(* IEC 61131-3 sources: daoli-st-library/DL_Device (part 37) *)

(* ---- FB_DL_WaferCassetteSlot.st ---- *)
(*==============================================================================
 * 组件名称 (Component)  : FB_DL_WaferCassetteSlot
 * 所属子库 (Sublibrary) : DL_Device
 * 当前版本 (Version)    : 1.0.0
 * 兼容性 (Platform)     : CODESYS 3.5 / TwinCAT 3 / 汇川 InoProShop（纯标准元素，零方言）
 * 功能描述 (Function)   : 花篮 25 槽占用双向计数与满/空判据。进片沿 +1、出片沿 −1，同拍
 *                         双沿按「物理不可能，必是抖动或逻辑错」双丢弃并报码；两个沿的净
 *                         额一次性施加，占用计数只有一处写入点；占用为 0 时的出片不借位到
 *                         25（借位会把满篮误判为空篮），锁存计数矛盾；位图按先低槽后高槽
 *                         顺序填充（顺序装片假设），出片清最低置位位。不做槽位光学检测、
 *                         不做花篮身份识别。
 * 溯源 (Origin)         : 道莅 clean-room 防御性实现
 * 本文件内含 (Contains) : TYPE E_DL_CassetteState / FUNCTION_BLOCK FB_DL_WaferCassetteSlot
 * 依赖 (Depends)        : 无（仅 Standard.library 的 SHL / SHR 与位运算）
 * 红线自检 (Redline)    : 无外部全局变量、无硬件地址直引 ｜ 全变量中英双语同行注释
 *                         槽数钳位 1~25 且写位图前判槽号 ｜ 占用计数单点写入（净额合并）
 *                         双沿沿实例无条件周期刷新 ｜ 枚举显式赋值 ｜ CASE 含 ELSE 兜底
 * 错误码表 (Codes)      : 16#0003_03B6 就绪（计数正常，含满/空稳态）
 *                         16#0003_03B7 故障级 清空请求在使能期被拒（清空须先失能）
 *                         16#0003_03B8 信息级 槽数 >25 已钳制（不置故障级标志）
 *                         16#0003_03B9 故障级 同拍进出双沿或满篮进片（请求双丢弃）
 *                         16#0003_03BA 故障级 空篮出片，锁存计数矛盾（不借位到 25）。
 *                                    本件 5 槽全用、无预留槽，已登记待裁定
 * 修订历史 (Revision)   : 2026-11-17  v1.0.0  首版入库 · R28 · 阶段三批 3
 * 验收向量 (Acceptance) : 正向 25 槽连续进满 → 占用 25、bFull、位图 16#01FF_FFFF；再出
 *                         1 片 → 占用 24、bFull=FALSE、16#0003_03B6
 *                         反向 空篮出片 → bCounterMismatch、占用保持 0、16#0003_03BA；
 *                         同拍进出双沿 → 16#0003_03B9 且双丢弃；槽数给 30 → 钳 25 +
 *                         16#0003_03B8（信息级）；使能期清空请求 → 16#0003_03B7 且不清
 *============================================================================*)

(*-----------------------------------------------------------------------------
 * 枚举: E_DL_CassetteState（归属本功能块，同文件发布，全库唯一定义）
 *----------------------------------------------------------------------------*)
TYPE E_DL_CassetteState :
(
    eEmpty := 0,    // 空篮：占用 0 / Empty cassette, no occupied slot
    ePart  := 10,   // 部分占用：0 < 占用 < 槽数 / Partially occupied
    eFull  := 20,   // 满篮：占用 = 槽数 / Full cassette
    eFault := 99    // 故障：计数矛盾锁存 / Fault, the counter contradiction is latched
);
END_TYPE

FUNCTION_BLOCK FB_DL_WaferCassetteSlot
VAR_INPUT
    bEnable      : BOOL := FALSE;         // 使能，FALSE 锁存位图（计数冻结） / Enable, FALSE freezes the slot map
    bLoadPulse   : BOOL := FALSE;         // 进片 +1，上升沿 / Load pulse, rising edge adds one
    bUnloadPulse : BOOL := FALSE;         // 出片 −1，上升沿 / Unload pulse, rising edge subtracts one
    bClear       : BOOL := FALSE;         // 清空（换花篮），须 bEnable=FALSE / Clear for a cassette change, requires bEnable FALSE
    uSlotCount   : UINT := 25;            // 槽数 [个]，域 1~25 / Slot count, domain 1 to 25
END_VAR
VAR_OUTPUT
    uOccupied    : UINT;                  // 占用槽数 [个] / Occupied slot count
    uEmptySlot   : UINT;                  // 空槽数 [个] / Empty slot count
    bFull        : BOOL;                  // 满篮判据 / Full criterion
    bEmpty       : BOOL;                  // 空篮判据 / Empty criterion
    uSlotMask    : DWORD;                 // 占用位图 bit0=第 1 槽 … bit24=第 25 槽 [bit]（25 位须 32 位容器，规格 WORD 无法表达） / Occupancy map, 25 bits need a 32-bit container
    bCounterMismatch : BOOL;              // 计数矛盾已锁存 / Counter contradiction latched
    eErr         : UDINT;                 // 错误码，段位 16#0003_xxxx / Error code in segment 16#0003_xxxx
END_VAR
VAR
    _eState      : E_DL_CassetteState := E_DL_CassetteState.eEmpty; // 占用状态 / Occupancy state
    _bInit       : BOOL := FALSE;         // 首扫标志，取非判定 / First-scan flag, tested negated
    _bMismatch   : BOOL := FALSE;         // 矛盾锁存状态量 / Contradiction latch state quantity
    _nNet        : INT;                   // 本拍净额（+进 −出） / Net delta of this scan
    _uSlotEff    : UINT := 25;            // 生效槽数（钳制后） / Effective slot count after clamping
    _uwOccupied  : UINT;                  // 占用内部唯一写点 / The single internal write point of the occupancy
    _rtrigLoad   : R_TRIG;                // 进片上升沿 / Rising edge of the load pulse
    _rtrigUnload : R_TRIG;                // 出片上升沿 / Rising edge of the unload pulse
END_VAR
VAR CONSTANT
    DL_CS_READY   : UDINT := 16#0003_03B6;  // 就绪码 / Ready code
    DL_CS_CLEAR_REJ : UDINT := 16#0003_03B7; // 故障级清空被拒码 / Fault code for a rejected clear request
    DL_CS_SLOT_CLAMP : UDINT := 16#0003_03B8; // 信息级槽数钳制码 / Info code for a clamped slot count
    DL_CS_BOTH    : UDINT := 16#0003_03B9;  // 故障级双沿或满篮进片码 / Fault code for double edges or a load on a full cassette
    DL_CS_UNDER   : UDINT := 16#0003_03BA;  // 故障级空篮出片码 / Fault code for an unload on an empty cassette
    DL_CS_SLOT_MAX : UINT := 25;            // 槽数上限 [个] / Slot count upper bound
    DL_CS_FULL_MASK : DWORD := 16#01FF_FFFF; // 25 槽满位图 [bit] / Full map of 25 slots
    DL_CS_BIT0      : DWORD := 16#0000_0001; // 位图零号位常量 [bit] / Bit zero constant of the map
END_VAR

// 段 1｜输出与单拍标志预置
eErr := 0;                                          // 错误码预清 / Error code pre-cleared
_nNet := 0;                                         // 净额预清 / Net delta pre-cleared

// 段 2｜双沿沿实例无条件周期刷新（R24：严禁置于分支内）
_rtrigLoad(CLK := bLoadPulse);                      // 进片沿 / Load edge
_rtrigUnload(CLK := bUnloadPulse);                  // 出片沿 / Unload edge

// 段 3｜首扫初始化（判据取非，R19）
IF NOT _bInit THEN
    _uwOccupied := 0;                               // 占用起点 0 [个] / Occupancy starts at zero
    _bInit := TRUE;                                 // 首扫只做一次 / The first scan runs once
END_IF

// 段 4｜槽数钳制（>25 钳制并报信息级；<1 钳制到 1）
IF uSlotCount > DL_CS_SLOT_MAX THEN
    _uSlotEff := DL_CS_SLOT_MAX;                    // 槽数上限钳制 [个] / Slot count clamped to the upper bound
    eErr := DL_CS_SLOT_CLAMP;                       // 信息级：槽数已钳制 / Info, the slot count was clamped
ELSIF uSlotCount < 1 THEN
    _uSlotEff := 1;                                 // 槽数下限钳制 [个] / Slot count clamped to the lower bound
    eErr := DL_CS_SLOT_CLAMP;                       // 信息级：槽数已钳制 / Info, the slot count was clamped
ELSE
    _uSlotEff := uSlotCount;                        // 采用组态槽数 [个] / Use the configured slot count
END_IF

// 段 5｜清空请求（须失能；使能期请求被拒并报码）
IF bClear THEN
    IF bEnable THEN
        eErr := DL_CS_CLEAR_REJ;                    // 故障级：使能期清空被拒 / Fault, a clear request while enabled is rejected
    ELSE
        _uwOccupied := 0;                           // 清空占用 [个] / Occupancy cleared
        _bMismatch := FALSE;                        // 矛盾锁存解除 / Contradiction latch released
        _eState := E_DL_CassetteState.eEmpty;       // 状态回空篮 / State back to empty
    END_IF
END_IF

// 段 6｜双向沿合并为净额（同拍双沿：物理不可能，双丢弃并报码）
IF _rtrigLoad.Q AND _rtrigUnload.Q THEN
    _nNet := 0;                                     // 双沿丢弃 / Both edges discarded
    eErr := DL_CS_BOTH;                             // 故障级：同拍双沿 / Fault, both edges in the same scan
ELSIF _rtrigLoad.Q THEN
    _nNet := 1;                                     // 进片 +1 / Load adds one
ELSIF _rtrigUnload.Q THEN
    _nNet := -1;                                    // 出片 −1 / Unload subtracts one
ELSE
    _nNet := 0;                                     // 无沿 / No edge
END_IF

// 段 7｜净额一次性施加（占用唯一写点；越界一律拒绝，不借位）
IF bEnable AND (NOT _bMismatch) THEN
    IF _nNet > 0 THEN
        IF _uwOccupied >= _uSlotEff THEN
            eErr := DL_CS_BOTH;                     // 故障级：满篮进片 / Fault, a load on a full cassette
        ELSE
            _uwOccupied := _uwOccupied + 1;         // 占用 +1（唯一写点）[个] / Occupancy incremented, the single write point
        END_IF
    ELSIF _nNet < 0 THEN
        IF _uwOccupied = 0 THEN
            _bMismatch := TRUE;                     // 空篮出片：锁存矛盾，不借位到 25 / Unload on an empty cassette, the contradiction is latched
            _eState := E_DL_CassetteState.eFault;
            eErr := DL_CS_UNDER;                    // 故障级：空篮出片 / Fault, an unload on an empty cassette
        ELSE
            _uwOccupied := _uwOccupied - 1;         // 占用 −1（唯一写点）[个] / Occupancy decremented, the single write point
        END_IF
    END_IF
END_IF

// 段 8｜位图维护（先低槽后高槽顺序填充；出片清最低置位位；写前判槽号 ≤ 槽数）
IF (NOT _bMismatch) AND (_uwOccupied > 0) THEN
    IF _uwOccupied >= DL_CS_SLOT_MAX THEN
        uSlotMask := DL_CS_FULL_MASK;               // 满 25 槽：满位图 [bit] / All 25 slots, the full map
    ELSE
        uSlotMask := SHL(DL_CS_BIT0, UINT_TO_UDINT(_uwOccupied)) - DL_CS_BIT0;   // 低 _uwOccupied 槽全置位 [bit] / The lowest occupied slots are set
    END_IF
ELSE
    uSlotMask := 16#0000_0000;                      // 空篮或矛盾锁存：位图清 / Empty or latched mismatch, the map is cleared
END_IF

// 段 9｜出口判据（占用/空槽/满/空）
uOccupied := _uwOccupied;                           // 占用出口 [个] / Occupancy output
IF _uwOccupied >= _uSlotEff THEN
    uEmptySlot := 0;                                // 满篮：空槽 0 [个] / Full, no empty slot
ELSE
    uEmptySlot := _uSlotEff - _uwOccupied;          // 空槽数 [个] / Empty slot count
END_IF
bFull := (_uwOccupied >= _uSlotEff);                // 满篮判据 / Full criterion
bEmpty := (_uwOccupied = 0);                        // 空篮判据 / Empty criterion
bCounterMismatch := _bMismatch;                     // 矛盾锁存出口 / Contradiction latch output

// 段 10｜占用状态映射（ENUM + CASE + ELSE 兜底）
CASE _eState OF
    E_DL_CassetteState.eEmpty:
        IF _uwOccupied > 0 THEN
            IF _uwOccupied >= _uSlotEff THEN
                _eState := E_DL_CassetteState.eFull;    // 直接满篮 / Straight to full
            ELSE
                _eState := E_DL_CassetteState.ePart;    // 部分占用 / Partially occupied
            END_IF
        END_IF
    E_DL_CassetteState.ePart:
        IF _uwOccupied = 0 THEN
            _eState := E_DL_CassetteState.eEmpty;       // 回空篮 / Back to empty
        ELSIF _uwOccupied >= _uSlotEff THEN
            _eState := E_DL_CassetteState.eFull;        // 转满篮 / To full
        END_IF
    E_DL_CassetteState.eFull:
        IF _uwOccupied = 0 THEN
            _eState := E_DL_CassetteState.eEmpty;       // 全出完回空篮 / Back to empty after unloading all
        ELSIF _uwOccupied < _uSlotEff THEN
            _eState := E_DL_CassetteState.ePart;        // 转部分占用 / To partially occupied
        END_IF
    E_DL_CassetteState.eFault:
        IF NOT _bMismatch THEN
            _eState := E_DL_CassetteState.eEmpty;       // 清空解除后回空篮 / Back to empty after the clear
        END_IF
    ELSE
        // 非法状态兜底：按矛盾锁存处理（安全侧）
        _bMismatch := TRUE;
        _eState := E_DL_CassetteState.eFault;
        eErr := DL_CS_UNDER;                            // 故障级：非法状态 / Fault, illegal state
END_CASE
IF eErr = 0 THEN
    eErr := DL_CS_READY;                                // 无事件回就绪码 / Ready code when nothing else applies
END_IF
END_FUNCTION_BLOCK

(* ---- FB_DL_WaferCoolChuck.st ---- *)
(*
  FB_DL_WaferCoolChuck  —  晶圆冷却吸盘（真空吸附确认 / 温控投运联锁 / 温度-真空双条件释放）/ Wafer cooling chuck
  分类 Category : DL_Device
  码位 Code     : 16#03_2_0B
  版本 Version  : 1.0.0
  来源 Source   : t2-2-lbp — IEC 61131-3 标准语义的道莅防御性实现
  溯源 Origin   : Lam LBP（背压冷却 / LBP 公开语义）借鉴，clean-room 实现，未复制任何源码行
  功能 Function : 1) 吸附链：发建立真空指令 → 真空度（负压绝对值）达 fVacConfirmKpa 且持续 tAttachConfirm
                     才确认 bClamped；确认后**才允许** bTempEnable（温控投运与吸附强联锁）；
                  2) 吸附失败按 nRetryMax 重试，每次重试重发建立指令，重试耗尽锁存 021B；
                  3) 释放链：须同时满足「温度 <= fTempAttachMaxC − 2 °C（回差）」与「真空已破」两条件，
                     任一不满足则不推进状态（温度不满足置 bInterlockBlocked，真空未破由 tReleaseTimeout 升级）；
                  4) 温度越限按「吸附中 / 未吸附」两路独立码归因（022B / 023B，R190 归因唯一）。
  边界 Boundary : ① fTempAttachMaxC 与环境上限 fAmbientMaxC 倒置（attach 上限 <= 环境上限）判组态错 020B，
                      状态进 eFault 且不投运；fVacConfirmKpa <= 0 / nRetryMax < 0 / 时间参数 <= 0 同判组态错；
                  ② **两路温度故障码不得共用**：吸附中越上限 = 022B（晶圆可能已吸附在超温盘面，必须锁存并
                      禁止再投温控）；未吸附时越上限 = 023B（只是盘面过温，允许冷却后继续）；
                  ③ 解除式自证：_bFault 清除 = rtReset.Q（引脚可满足）；022B / 023B 另可由
                      「温度回落至 fTempAttachMaxC − DL_TEMP_HYST_C 以下」按码专清（R188 可达清除边）；
                  ④ 释放期真空未破不推进状态（不靠延时硬推），由 tReleaseTimeout 升级为 024B 锁存；
                  ⑤ 注入件故障（iVac.bFault / iTempZone.bFault）→ 拒绝新吸附并置信息级 013B（不置 bError，
                      故障属主是被注入件，本件只用其 uErrorId 做归因透出）；
                  ⑥ bTempEnable 仅在 eClamped / eCooling 两相为真，其余相（含 eReleasing / eFault）恒 FALSE。
  依赖 Depends  : I_DL_VacuumGenerator（DL_Device 既有契约）、I_DL_TemperatureZone（DL_Device 既有契约）；
                  仅 Standard.library（TON / R_TRIG / ABS / MIN / MAX），接口只注入不实例化
  同拍双窗配比  : tAttachConfirm（吸附确认驻留）与 tReleaseTimeout（释放超时）不同源；配比约束
                  tAttachConfirm <= tReleaseTimeout，避免释放判据比吸附确认更早失效（R100）

  码表 Error codes（本件格 03_2_0B，子码步进 +0x10）:
    16#0003_020B 故障级：组态非法（温度上限倒置 / 真空确认门限 <= 0 / 重试次数 < 0 / 时间参数 <= 0）
    16#0003_021B 故障级：吸附失败且重试耗尽（真空未达 fVacConfirmKpa，锁存）
    16#0003_022B 故障级：吸附保持中盘面温度越上限（禁止再投温控，锁存）
    16#0003_023B 故障级：未吸附状态下盘面温度越上限（盘面过温，冷却后可解）
    16#0003_024B 故障级：释放超时（tReleaseTimeout 到点真空仍未破，锁存）
    16#0003_025B 故障级：状态机落 ELSE 兜底（非法相位 ID）
    16#0003_010B 信息级：释放被温度联锁阻断（温度未回落到允许上限以下，不置 bError）
    16#0003_011B 信息级：吸附确认完成（bClamped 上升拍，不置 bError）
    16#0003_012B 信息级：吸附重试一次（本次未达真空门限，重发建立指令）
    16#0003_013B 信息级：注入件故障，拒绝吸附（iVac.bFault 或 iTempZone.bFault，不置 bError）

  修订历史 Revision :
    2026-11-18  v1.0.0  R37 首版
*)

TYPE E_DL_ChuckState :
(
    eIdle       := 0,   // 空闲：未吸附、温控断开 / Idle, no clamping, temperature control off
    eEvacuating := 10,  // 吸附中：建立真空并等待确认 / Evacuating, waiting for the vacuum confirmation
    eClamped    := 20,  // 已吸附：真空确认，温控待投运 / Clamped, vacuum confirmed, temperature control pending
    eCooling    := 30,  // 冷却中：温控已投运并保持 / Cooling, temperature control commissioned and holding
    eReleasing  := 40,  // 释放中：破真空，等温度与真空双条件 / Releasing, awaiting both temperature and vacuum release
    eFault      := 90   // 故障：锁存待复位（温度回落或复位沿）/ Fault, latched until reset or temperature recovery
);
END_TYPE

FUNCTION_BLOCK FB_DL_WaferCoolChuck
VAR_INPUT
    bEnable      : BOOL := FALSE;              // 总使能，FALSE 时断温控并停吸附 / Master enable, low level cuts the temperature control
    bReset       : BOOL := FALSE;              // 复位，上升沿清故障锁存 / Reset, rising edge clears the latch
    bClampCmd    : BOOL := FALSE;              // 吸附命令（电平，上升沿受理）/ Clamp command, accepted on a rising edge
    bReleaseCmd  : BOOL := FALSE;              // 释放命令（电平，上升沿受理）/ Release command, accepted on a rising edge
    fTempAttachMaxC : REAL := 45.0;            // 脱附允许温度上限 [°C]，域 > fAmbientMaxC / Maximum temperature permitting a release [degC]
    fAmbientMaxC : REAL := 25.0;               // 环境温度上限 [°C]，组态交叉校验用 / Ambient ceiling used by the configuration cross-check [degC]
    fVacConfirmKpa  : REAL := 60.0;            // 真空确认门限（负压绝对值）[kPa]，域 > 0 / Vacuum confirmation threshold, magnitude [kPa]
    fVacBreakKpa : REAL := 5.0;                // 判破真空门限（负压绝对值）[kPa]，域 > 0 / Vacuum-broken threshold, magnitude [kPa]
    tAttachConfirm : TIME := T#300MS;          // 吸附确认驻留时间 [ms]，域 > 0 / Attachment confirm dwell [ms]
    tRetryTimeout : TIME := T#2S;              // 单次吸附等待上限 [ms]，超时即重试 / Per-attempt vacuum budget [ms]
    tReleaseTimeout : TIME := T#5S;            // 释放超时 [ms]，超时升级故障 / Release timeout before raising a fault [ms]
    nRetryMax    : INT := 3;                   // 最大重试次数 [次]，域 >= 0 / Maximum retry count
    fCoolSetpointC : REAL := 20.0;             // 冷却设定温度 [°C]，投运时下发 / Cooling setpoint pushed on commissioning [degC]
END_VAR
VAR_OUTPUT
    bClamped     : BOOL;                       // 已吸附（真空确认）标志 / Clamped flag, vacuum confirmed
    bTempEnable  : BOOL;                       // 温控投运命令（吸附确认后才为真）/ Temperature control enable, true only while clamped
    bInterlockBlocked : BOOL;                  // 联锁阻断标志（释放被温度条件挡住）/ Interlock blocked, the release is held by temperature
    fVacKpa      : REAL;                       // 真空度（负压绝对值）[kPa]，诊断用 / Vacuum magnitude [kPa] for diagnostics
    fTempC       : REAL;                       // 盘面实测温度 [°C] / Chuck temperature [degC]
    nRetryCount  : INT;                        // 已重试次数 [次] / Retry counter
    bValid       : BOOL;                       // 判据可用标志 / Criteria usable
    bError       : BOOL;                       // 故障标志，派生自锁存 / Fault flag derived from the latch
    nErrId       : UDINT;                      // 事件码，0 = 无事件 / Event code, 0 = no event
    eStateOut    : E_DL_ChuckState;            // 状态出口，段尾单点映射 / State outlet, mapped at the tail
END_VAR
VAR_IN_OUT
    iVac         : I_DL_VacuumGenerator;       // 真空发生器接口引用（注入，不实例化）/ Vacuum generator reference, injected
    iTempZone    : I_DL_TemperatureZone;       // 温控区接口引用（注入，不实例化）/ Temperature zone reference, injected
END_VAR
VAR
    tonAttach    : TON;                        // 吸附确认驻留计时，每拍无条件调用 / Attachment confirm timer, called unconditionally
    tonAttempt   : TON;                        // 单次吸附等待计时，每拍无条件调用 / Per-attempt budget timer, called unconditionally
    tonRelease   : TON;                        // 释放超时计时，每拍无条件调用 / Release timeout timer, called unconditionally
    tonHeart     : TON;                        // 周期心跳窗，自复位 / Periodic heartbeat window, self-resetting
    rtReset      : R_TRIG;                     // 复位上升沿 / Reset rising edge
    rtClamp      : R_TRIG;                     // 吸附命令上升沿 / Clamp command rising edge
    rtRelease    : R_TRIG;                     // 释放命令上升沿 / Release command rising edge
    _eState      : E_DL_ChuckState := E_DL_ChuckState.eIdle;  // 内部相位（CASE 唯一写入目标）/ Internal phase
    _uFault      : UDINT;                      // 故障码锁存 / Latched fault code
    _uInfo       : UDINT;                      // 信息码，每拍重算 / Information code, recomputed per scan
    _bFault      : BOOL;                       // 故障锁存位 / Latched fault bit
    _bParamBad   : BOOL;                       // 组态非法聚合 / Configuration invalid aggregate
    _bVacOk      : BOOL;                       // 真空达确认门限 / Vacuum reached the confirm threshold
    _bVacBroken  : BOOL;                       // 真空已破 / Vacuum broken
    _bTempHigh   : BOOL;                       // 温度越脱附允许上限 / Temperature above the release limit
    _bTempOkRel  : BOOL;                       // 温度满足释放条件（带回差）/ Temperature satisfies the release with hysteresis
    _bInjectFault: BOOL;                       // 注入件故障 / An injected component reports a fault
    _bCmdEvac    : BOOL;                       // 建立真空单发请求（段 6 落地）/ One-shot evacuate request, applied in segment 6
    _bCmdBlow    : BOOL;                       // 破真空单发请求（段 6 落地）/ One-shot blow-off request, applied in segment 6
    _bCmdStop    : BOOL;                       // 双阀全断单发请求（段 6 落地）/ One-shot stop request, applied in segment 6
    _bTempSet    : BOOL;                       // 下发设定温度单发请求 / One-shot setpoint request
    _bTempOn     : BOOL;                       // 温控投运单发请求 / One-shot temperature commission request
    _bTempOff    : BOOL;                       // 温控断电单发请求 / One-shot temperature decommission request
    _bClampedPrev: BOOL;                       // 上拍吸附快照 / Previous-scan clamped snapshot
    _bHeartBreak : BOOL := TRUE;               // 心跳窗断输入一拍 / One-scan heartbeat break
    _nRetry      : INT;                        // 重试计数保持量 [次] / Held retry counter
    _bAttemptBrk : BOOL := TRUE;               // 单次等待计时断输入一拍 / One-scan budget break
    _bRelBreak   : BOOL := TRUE;               // 释放超时计时断输入一拍 / One-scan release break
END_VAR
VAR CONSTANT
    DL_TEMP_HYST_C : REAL := 2.0;      // 释放温度回差 [°C]（规格固定 2 °C）/ Release temperature hysteresis, fixed at two degrees
    DL_EPS         : REAL := 1.0E-6;   // 判零容差 [1] / Zero tolerance
    DL_HEART_WINDOW : TIME := T#2S;    // 心跳观察窗 [ms]，自复位节拍 / Heartbeat window, self-resetting
    DL_VAL_LIM_C   : REAL := 500.0;    // 温度有限性上限 [°C] / Temperature magnitude ceiling [degC]
    DL_VAL_LIM_KPA : REAL := 200.0;    // 真空有限性上限 [kPa] / Vacuum magnitude ceiling [kPa]
END_VAR

(* —— 段 0：定时器与边缘检测无条件周期刷新（R182：调用语句不得置于 IF / CASE 内） —— *)
rtReset(CLK := bReset);                                        // 复位上升沿，每拍必调
rtClamp(CLK := bClampCmd);                                     // 吸附命令上升沿，每拍必调
rtRelease(CLK := bReleaseCmd);                                 // 释放命令上升沿，每拍必调
tonHeart(IN := (NOT tonHeart.Q) AND (NOT _bHeartBreak), PT := DL_HEART_WINDOW);  // 心跳窗自复位
_bHeartBreak := FALSE;                                         // 断输入拍在调用后自清
tonAttach(IN := (_eState = E_DL_ChuckState.eEvacuating) AND _bVacOk, PT := tAttachConfirm);  // 吸附确认驻留
tonAttempt(IN := (_eState = E_DL_ChuckState.eEvacuating) AND (NOT _bVacOk) AND (NOT _bAttemptBrk),
           PT := tRetryTimeout);                               // 单次等待（表达式入参）
_bAttemptBrk := FALSE;                                         // 断输入拍在调用后自清
tonRelease(IN := (_eState = E_DL_ChuckState.eReleasing) AND (NOT _bVacBroken) AND (NOT _bRelBreak),
           PT := tReleaseTimeout);                             // 释放超时（表达式入参）
_bRelBreak := FALSE;                                           // 断输入拍在调用后自清

(* —— 段 1：单拍量预清零（计数 / 保持量 / 锁存不入清单，R187①） —— *)
_uInfo        := 16#0000_0000;   // 信息码每拍重算
bError        := FALSE;          // 故障出口每拍重算，段 7 由锁存派生
bValid        := FALSE;          // 可用标志缺省 FALSE
bClamped      := FALSE;          // 吸附出口缺省 FALSE，段 8 单点置位
bTempEnable   := FALSE;          // 温控投运缺省 FALSE（失能优先）
bInterlockBlocked := FALSE;      // 联锁阻断缺省 FALSE
_bParamBad    := FALSE;          // 组态非法预清零
_bVacOk       := FALSE;          // 真空确认判据预清零
_bVacBroken   := FALSE;          // 破真空判据预清零
_bTempHigh    := FALSE;          // 温度越限判据预清零
_bTempOkRel   := FALSE;          // 释放温度条件预清零
_bInjectFault := FALSE;          // 注入件故障预清零
_bCmdEvac     := FALSE;          // 单发请求预清零（本次 CASE 可重新置位）
_bCmdBlow     := FALSE;          // 破真空请求预清零
_bCmdStop     := FALSE;          // 全断请求预清零
_bTempSet     := FALSE;          // 设温请求预清零
_bTempOn      := FALSE;          // 投运请求预清零
_bTempOff     := FALSE;          // 断电请求预清零

(* —— 段 2：复位沿清锁存（按码专清 / 恢复沿清码两路径互不掩盖，R188） —— *)
IF rtReset.Q THEN
    _bFault := FALSE;            // 复位沿清锁存位
    _uFault := 16#0000_0000;     // 复位沿清锁存码
    _nRetry := 0;                // 复位沿清重试计数（吸附链重新起算）
    _uInfo  := 16#0000_0000;     // 复位拍不报旧信息
END_IF

(* —— 段 3：组态域闸 + 输入有限性（覆盖全部参与判据换算的引脚，R151） —— *)
IF (fTempAttachMaxC <> fTempAttachMaxC) OR (fTempAttachMaxC > DL_VAL_LIM_C) OR
   (fTempAttachMaxC <= fAmbientMaxC) THEN
    _bParamBad := TRUE;          // 脱附允许上限非法或与环境上限倒置（上限须高于环境）
END_IF
IF (fVacConfirmKpa <> fVacConfirmKpa) OR (fVacConfirmKpa <= 0.0) OR (fVacConfirmKpa > DL_VAL_LIM_KPA) THEN
    _bParamBad := TRUE;          // 真空确认门限非法（确认判据的分母语义）
END_IF
IF (fVacBreakKpa <> fVacBreakKpa) OR (fVacBreakKpa <= 0.0) OR (fVacBreakKpa >= fVacConfirmKpa) THEN
    _bParamBad := TRUE;          // 破真空门限非法或与确认门限倒置（会形成永判未破的死区）
END_IF
IF (fCoolSetpointC <> fCoolSetpointC) OR (fCoolSetpointC <= fAmbientMaxC) THEN
    _bParamBad := TRUE;          // 冷却设定非法（须高于环境上限，否则只在环境温度上打转）
END_IF
IF nRetryMax < 0 THEN
    _bParamBad := TRUE;          // 重试次数为负非法
END_IF
IF (TIME_TO_DINT(tAttachConfirm) <= 0) OR (TIME_TO_DINT(tRetryTimeout) <= 0) OR
   (TIME_TO_DINT(tReleaseTimeout) <= 0) THEN
    _bParamBad := TRUE;          // 三个时间参数均须 > 0
END_IF
IF _bParamBad THEN
    _uFault := 16#0003_020B;     // 故障级：组态非法
    _bFault := TRUE;             // 锁存位置位（复位沿可清）
    bError  := TRUE;             // 故障标志置位（R45 配对）
    _eState := E_DL_ChuckState.eFault;  // 进故障相
END_IF

(* —— 段 4：反馈采集与判据（只读属性，零命令下发） —— *)
fVacKpa := ABS(iVac.fPressure);                 // 真空度 = 负压绝对值 [kPa]
fTempC  := iTempZone.fTempActual;               // 盘面实测温度 [°C]
IF (fVacKpa <> fVacKpa) OR (fVacKpa > DL_VAL_LIM_KPA) THEN
    _bParamBad := TRUE;                         // 真空反馈非有限或超上界：判输入异常（不得静默当作无真空）
    _uFault := 16#0003_020B;                    // 故障级：输入异常归入组态/输入异常码
    _bFault := TRUE;                            // 锁存
    bError  := TRUE;                            // 故障标志置位（R45 配对）
    _eState := E_DL_ChuckState.eFault;          // 进故障相
END_IF
_bVacOk      := (fVacKpa >= fVacConfirmKpa);    // 达确认门限
_bVacBroken  := (fVacKpa <= fVacBreakKpa);      // 已破真空（门限带迟滞，两门限已证不倒置）
_bTempHigh   := (fTempC > fTempAttachMaxC);     // 越脱附允许上限
_bTempOkRel  := (fTempC <= (fTempAttachMaxC - DL_TEMP_HYST_C));  // 释放条件：回落 2 °C（回差）
_bInjectFault := iVac.bFault OR iTempZone.bFault;                // 注入件故障聚合

(* —— 段 5：温度越限两路归因（吸附中 / 未吸附，码不共用，R190） —— *)
IF (fTempC < -DL_VAL_LIM_C) OR (fTempC > DL_VAL_LIM_C) THEN
    _bParamBad := TRUE;                          // 温度非有限：按组态/输入异常处理，不伪造越限
    _uFault := 16#0003_020B;                     // 故障级：输入非有限归入组态/输入异常码
    _bFault := TRUE;                             // 锁存
    bError  := TRUE;                             // 故障标志置位（R45 配对）
    _eState := E_DL_ChuckState.eFault;           // 进故障相
ELSIF _bTempHigh THEN
    IF (_eState = E_DL_ChuckState.eClamped) OR (_eState = E_DL_ChuckState.eCooling) THEN
        _uFault := 16#0003_022B;                 // 故障级：吸附保持中温度越上限（独立码）
        _bFault := TRUE;                         // 锁存
        bError  := TRUE;                         // 故障标志置位（R45 配对）
        _eState := E_DL_ChuckState.eFault;       // 进故障相（温控强制断）
    ELSE
        _uFault := 16#0003_023B;                 // 故障级：未吸附状态下盘面过温（独立码，冷却后可解）
        _bFault := TRUE;                         // 锁存
        bError  := TRUE;                         // 故障标志置位（R45 配对）
        _eState := E_DL_ChuckState.eFault;       // 进故障相
    END_IF
END_IF
IF (_uFault = 16#0003_022B) OR (_uFault = 16#0003_023B) THEN
    IF _bTempOkRel THEN
        _uFault := 16#0000_0000;                 // 按码专清：温度回落至回差带以下 → 温度类故障可解
        _bFault := FALSE;                        // 锁存位同步清（复位沿路径互不掩盖）
    END_IF
END_IF

(* —— 段 6：相位机（只做迁移与单发请求置位；命令下发在本段末统一执行） —— *)
CASE _eState OF

E_DL_ChuckState.eIdle:
    _nRetry := 0;                                            // 空闲：重试计数归零（唯一清零点在本相）
    IF rtClamp.Q THEN
        IF (NOT bEnable) OR _bInjectFault THEN
            _uInfo := 16#0003_013B;                          // 信息级：注入件故障或未使能，拒绝吸附
        ELSIF _bFault THEN
            _uInfo := 16#0003_013B;                          // 信息级：存在未复位故障，拒绝吸附
        ELSE
            _eState := E_DL_ChuckState.eEvacuating;          // 进吸附相
            _bCmdEvac := TRUE;                               // 首个建立真空指令（单发）
            _bAttemptBrk := TRUE;                            // 单次等待计时从零开始
        END_IF
    END_IF

E_DL_ChuckState.eEvacuating:
    IF (NOT bEnable) OR _bInjectFault THEN
        _bCmdStop := TRUE;                                   // 全断双阀（安全侧），退出吸附
        _uInfo := 16#0003_013B;                              // 信息级：注入件故障，中止吸附
        _eState := E_DL_ChuckState.eIdle;                    // 回空闲
    ELSIF tonAttach.Q THEN
        _eState := E_DL_ChuckState.eClamped;                 // 吸附确认：真空达标并驻留完成
        _nRetry := 0;                                        // 确认成功：重试计数归零
        _uInfo  := 16#0003_011B;                             // 信息级：吸附确认完成
        _bTempSet := TRUE;                                   // 下发冷却设定温度（单发）
    ELSIF tonAttempt.Q THEN
        IF _nRetry < nRetryMax THEN
            _nRetry := _nRetry + 1;                          // 重试计数 +1
            _bCmdEvac := TRUE;                               // 重发建立真空指令（单发）
            _bAttemptBrk := TRUE;                            // 单次等待计时重启
            _uInfo := 16#0003_012B;                          // 信息级：吸附重试一次
        ELSE
            _uFault := 16#0003_021B;                         // 故障级：重试耗尽，吸附失败锁存
            _bFault := TRUE;                                 // 锁存
            bError  := TRUE;                                 // 故障标志置位（R45 配对）
            _bCmdStop := TRUE;                               // 全断双阀（不在失败态继续抽气）
            _eState := E_DL_ChuckState.eFault;               // 进故障相
        END_IF
    ELSIF rtRelease.Q THEN
        _bCmdStop := TRUE;                                   // 吸附未确认即释放：全断双阀
        _eState := E_DL_ChuckState.eIdle;                    // 回空闲（真空未建立，无需破真空）
    END_IF

E_DL_ChuckState.eClamped:
    _bTempOn := TRUE;                                        // 已吸附：允许投运温控（本相唯一置位点）
    IF (NOT bEnable) OR _bInjectFault THEN
        _bTempOff := TRUE;                                   // 断温控
        _bCmdStop := TRUE;                                   // 全断双阀（保守：失能即解除吸附保持）
        _uInfo := 16#0003_013B;                              // 信息级：注入件故障或失能
        _eState := E_DL_ChuckState.eIdle;                    // 回空闲
    ELSIF rtRelease.Q THEN
        _eState := E_DL_ChuckState.eReleasing;               // 进释放相（温度与真空双条件在相内判）
        _bRelBreak := TRUE;                                  // 释放超时计时从零开始
        _bCmdBlow := TRUE;                                   // 破真空指令（单发）
    ELSE
        _eState := E_DL_ChuckState.eCooling;                 // 确认后进冷却保持相
    END_IF

E_DL_ChuckState.eCooling:
    _bTempOn := TRUE;                                        // 冷却中：温控保持投运
    IF (NOT bEnable) OR _bInjectFault THEN
        _bTempOff := TRUE;                                   // 断温控
        _bCmdStop := TRUE;                                   // 全断双阀
        _uInfo := 16#0003_013B;                              // 信息级：注入件故障或失能
        _eState := E_DL_ChuckState.eIdle;                    // 回空闲
    ELSIF rtRelease.Q THEN
        _eState := E_DL_ChuckState.eReleasing;               // 进释放相
        _bRelBreak := TRUE;                                  // 释放超时计时从零开始
        _bCmdBlow := TRUE;                                   // 破真空指令（单发）
    END_IF

E_DL_ChuckState.eReleasing:
    IF _bVacBroken AND _bTempOkRel THEN
        _bTempOff := TRUE;                                   // 温控断电（释放完成，不再控温）
        _eState := E_DL_ChuckState.eIdle;                    // 双条件成立：回空闲
    ELSIF NOT _bTempOkRel THEN
        bInterlockBlocked := TRUE;                           // 温度未回落：联锁阻断，**状态不推进**
        _uInfo := 16#0003_010B;                              // 信息级：释放被温度联锁阻断
        IF tonRelease.Q THEN
            _uFault := 16#0003_024B;                         // 故障级：释放超时（温度与真空双失败）
            _bFault := TRUE;                                 // 锁存
            bError  := TRUE;                                 // 故障标志置位（R45 配对）
            _eState := E_DL_ChuckState.eFault;               // 进故障相
        END_IF
    ELSIF tonRelease.Q THEN
        _uFault := 16#0003_024B;                             // 故障级：真空未破且超时（真空侧失败）
        _bFault := TRUE;                                     // 锁存
        bError  := TRUE;                                     // 故障标志置位（R45 配对）
        _eState := E_DL_ChuckState.eFault;                   // 进故障相
    END_IF

E_DL_ChuckState.eFault:
    _bTempOff := TRUE;                                       // 故障：温控强制断电（安全侧）
    _bCmdStop := TRUE;                                       // 故障：双阀全断（保持现状，不主动吹气）
    IF (NOT _bFault) AND (NOT _bParamBad) AND bEnable THEN
        _eState := E_DL_ChuckState.eIdle;                    // 锁存已清且组态合法：回空闲
    END_IF

ELSE
    _uFault := 16#0003_025B;                                 // 故障级：相位 ID 越界（枚举兜底）
    _bFault := TRUE;                                         // 锁存
    bError  := TRUE;                                         // 故障标志置位（R45 配对）
    _eState := E_DL_ChuckState.eFault;                       // 强制回故障相
END_CASE

(* —— 段 6A：单发命令落地（每拍最多一次，禁在 CASE 内直呼接口方法） —— *)
_bTempOn  := _bTempOn  AND (NOT _bFault);   // 故障期不投运温控（门控挂状态量）
_bTempSet := _bTempSet AND (NOT _bFault);   // 故障期不下发设定
IF _bCmdEvac THEN
    _bCmdEvac := FALSE;                     // 先清标志再下发，防方法内异常导致重复调用
    _bCmdEvac := iVac.CmdEvacuate();        // 建立真空（返回受理结果，未受理则由重试链兜底）
END_IF
IF _bCmdBlow THEN
    _bCmdBlow := FALSE;                     // 先清标志
    _bCmdBlow := iVac.CmdBlowOff();         // 破真空（实现块输出定宽脉冲）
END_IF
IF _bCmdStop THEN
    _bCmdStop := FALSE;                     // 先清标志
    _bCmdStop := iVac.CmdStop();            // 双阀全断（保持现状）
END_IF
IF _bTempSet THEN
    _bTempSet := FALSE;                     // 先清标志
    _bTempSet := iTempZone.SetSetpoint(fTemp := fCoolSetpointC);  // 下发冷却设定
END_IF
IF _bTempOn THEN
    _bTempOn := FALSE;                      // 先清标志
    iTempZone.CmdEnable(bOn := TRUE);       // 温控投运（无返回，靠反馈确认）
END_IF
IF _bTempOff THEN
    _bTempOff := FALSE;                     // 先清标志
    iTempZone.CmdEnable(bOn := FALSE);      // 温控断电（无返回，安全侧动作）
END_IF

(* —— 段 7：故障码优先级链（每个 bError 置位源在此均有码，R45 配对） —— *)
IF _bParamBad THEN
    bError := TRUE;                         // 组态非法：码已在段 3/段 5 置位（020B），此处仅保证配对
END_IF

(* —— 段 8：出口单点映射（名实同源；锁存码回放，禁同拍抹除） —— *)
bClamped := (_eState = E_DL_ChuckState.eClamped) OR (_eState = E_DL_ChuckState.eCooling);  // 吸附保持出口
bTempEnable := bClamped AND bEnable AND (NOT _bFault);   // 温控投运：仅吸附保持且无故障且使能
nRetryCount := _nRetry;                                  // 重试计数出口
eStateOut   := _eState;                                  // 状态出口
IF _bFault THEN
    nErrId := _uFault;                                   // 故障锁存码回放（不在故障相按当下输入重推）
    bError := TRUE;                                      // 故障出口派生自锁存
ELSE
    nErrId := _uInfo;                                    // 信息码
END_IF
bValid := bEnable AND (NOT _bFault) AND (NOT _bParamBad);  // 判据可用

END_FUNCTION_BLOCK

(* ---- FB_DL_WaferHandoffSeq.st ---- *)
(*==============================================================================
 * 组件名称 (Component)  : FB_DL_WaferHandoffSeq
 * 所属子库 (Sublibrary) : DL_Device
 * 前缀     (Prefix)     : FB_DL_
 * 当前版本 (Version)    : 1.0.0
 * 兼容性   (Platform)   : CODESYS 3.5 / TwinCAT 3 / 汇川 InoProShop / Schneider
 *                         Machine Expert；纯 IEC 61131-3（第 3 版），
 *                         仅依赖标准库 TON / R_TRIG，零厂商方言
 * 作者     (Author)     : 道莅代码库 · PLC编程专家（R31）
 * 开源溯源 (Origin)     : 双机械手晶圆交接防碰撞握手公开工艺语义（行业池），
 *                         道莅 clean-room 防御性实现，未复制任何外部源码行
 * 功能描述 (Function)   : 双机械手交接防碰撞握手顺控件。步序：A/B 就位 →
 *                         A 释放 → B 吸持 → A 撤离 → B 撤离 → 完成。
 *                         互斥核心写死：任一方未撤离交接区，另一方不得获得
 *                         移动放行；防碰撞为安全侧语义。双请求同拍按固定
 *                         优先 A 先（头注释留档）。到位信号非预期跳变
 *                         即中止锁故障。不套通用 InterlockMatrix（判定段
 *                         与执行段不共享状态机教训，本件自带专用互锁）。
 * 状态机   (States)     : eIdle 待机 / eMoveAIn A 进场 / eMoveBIn B 进场 /
 *                         eARelease A 释放 / eWaitGripB B 吸持确认 /
 *                         eAExit A 撤离 / eBExit B 撤离 / eDone 单拍完成 /
 *                         eFault 故障锁定（CASE 带 ELSE 兜底）。
 * 码位     (Codes)      : 16#0003_03F2 信息级：双请求同拍（A 优先留档，
 *                                      不置 bError）
 *                         16#0003_03F3 故障级：步超时
 *                         16#0003_03F4 故障级：移动互锁违例（防御断言）
 *                         16#0003_03F5 故障级：到位/吸持反馈矛盾（非预期跳变）
 *                         16#0003_03F6 故障级：状态非法（ELSE 兜底）
 * 边界防错 (Boundary)   : 1 移动放行由状态机逐拍重算派生，非锁存量；
 *                         2 步超时 TON 按步断输入（步切换拍单拍断输入）；
 *                         3 TON/R_TRIG 实例每拍无条件刷新；
 *                         4 故障锁存可达解除路径：撤使能（bEn 下降）回待机清码；
 *                         5 bDone 为单拍脉冲（R27 跨拍须清零）。
 * 修订历史 (Revision)   : 2026-11-18 v1.0.0 首版入库（R31 · 阶段三 · 序 9）
 *==============================================================================*)

(*------------------------------------------------------------------------------
 * 枚举: E_DL_HandoffStep（归属本功能块，同文件发布，全库唯一属主）
 *----------------------------------------------------------------------------*)
TYPE E_DL_HandoffStep :
(
    eIdle      := 0,    // 待机：等待双方请求 / Idle, waiting for both requests
    eMoveAIn   := 10,   // A 进场：放行 A 至就位 / A entering, move permit to A
    eMoveBIn   := 20,   // B 进场：放行 B 至就位 / B entering, move permit to B
    eARelease  := 30,   // A 释放：等待 A 吸持反馈消失 / A releasing, wait grip-A drop
    eWaitGripB := 40,   // B 吸持：等待 B 吸持确认 / B gripping, wait grip-B confirm
    eAExit     := 50,   // A 撤离：放行 A 至出场 / A exiting, move permit to A
    eBExit     := 60,   // B 撤离：放行 B 至出场 / B exiting, move permit to B
    eDone      := 70,   // 完成：单拍脉冲后回待机 / Done, one-scan pulse then idle
    eFault     := 99    // 故障：锁定等待撤使能复位 / Fault, latched until disabled
);
END_TYPE

(*==============================================================================
 * 功能块: FB_DL_WaferHandoffSeq
 * 调用约定: 每个扫描周期无条件调用一次；bMoveA/bMoveB 为移动放行指令。
 *==============================================================================*)
FUNCTION_BLOCK FB_DL_WaferHandoffSeq
VAR_INPUT
    bReqA    : BOOL := FALSE;         // 机械手 A 交接请求 / Robot A handoff request
    bReqB    : BOOL := FALSE;         // 机械手 B 交接请求 / Robot B handoff request
    bPosA    : BOOL := FALSE;         // A 交接区就位反馈 / Robot A in-position feedback
    bPosB    : BOOL := FALSE;         // B 交接区就位反馈 / Robot B in-position feedback
    bGripA   : BOOL := FALSE;         // A 吸持反馈 / Robot A grip feedback
    bGripB   : BOOL := FALSE;         // B 吸持反馈 / Robot B grip feedback
    bEn      : BOOL := FALSE;         // 使能，下降沿为故障可达解除路径 / Enable, falling edge is fault release path
    tStep    : TIME := T#5S;          // 单步超时 [毫秒] / Per-step timeout [ms]
END_VAR
VAR_OUTPUT
    eStep    : E_DL_HandoffStep;      // 当前步状态 / Current handshake step
    bMoveA   : BOOL;                  // A 移动放行（互锁派生）/ Robot A move permit, interlocked
    bMoveB   : BOOL;                  // B 移动放行（互锁派生）/ Robot B move permit, interlocked
    bDone    : BOOL;                  // 交接完成单拍脉冲（R27）/ Handoff done one-scan pulse
    bError   : BOOL;                  // 故障标志，与故障级码配对（R45）/ Fault flag paired with fault codes
    uErrorId : UDINT;                 // 错误码，0 = 无错 / Error code, 0 = none
END_VAR
VAR
    tonStep  : TON;                   // 步超时定时器，每拍无条件刷新 / Step timeout timer, refreshed every scan
    rTrigA   : R_TRIG;                // A 请求沿检测，每拍无条件刷新 / Request-A edge detector
    rTrigB   : R_TRIG;                // B 请求沿检测，每拍无条件刷新 / Request-B edge detector
    eStatePrev : E_DL_HandoffStep;    // 上一拍步快照 / Previous step snapshot
    bStepRst : BOOL;                  // 步切换拍单拍断超时输入 / One-scan timeout input break on step change
    uInfoOne : UDINT;                 // 信息级单拍码暂存 / One-scan info code staging
    uCodeLatch : UDINT;               // 故障级锁存码 / Latched fault code
    bInit    : BOOL := TRUE;          // 首扫标志 / First-scan flag
END_VAR
VAR CONSTANT
    DL_WHS_ZERO : UDINT := 16#0000_0000; // 零码常量 / Zero code constant
END_VAR

// ---- 段 1｜边沿与定时器实例无条件周期刷新（红线：禁入条件分支）----------------
rTrigA(CLK := bReqA);                                 // A 请求沿检测 / Request-A edge detection
rTrigB(CLK := bReqB);                                 // B 请求沿检测 / Request-B edge detection
tonStep(IN := (eStep <> eIdle) AND (eStep <> eDone) AND (eStep <> eFault)
        AND (NOT bStepRst), PT := tStep);             // 步超时计时，步切换拍断输入 / Step timing, broken on step change

// ---- 段 2｜步切换检测（供超时按步断输入）----------------------------------------
bStepRst := (eStep <> eStatePrev) OR bInit;           // 步变化即断输入 / Step change breaks timing input
eStatePrev := eStep;                                  // 快照留痕 / Snapshot previous step
bInit := FALSE;                                       // 清首扫标志 / Clear first-scan flag

// ---- 段 3｜移动放行派生：互斥核心，任一方未撤离另一方不得放行 --------------------
bMoveA := (eStep = eMoveAIn) OR (eStep = eAExit);     // A 放行仅进场/撤离步 / A permit only in enter/exit steps
bMoveB := (eStep = eMoveBIn) OR (eStep = eBExit);     // B 放行仅进场/撤离步 / B permit only in enter/exit steps

// ---- 段 4｜状态机（CASE 带 ELSE 兜底锁故障）--------------------------------------
CASE eStep OF
    eIdle:
        bDone := FALSE;                               // 待机清完成脉冲 / Idle clears done pulse
        IF bEn AND rTrigA.Q AND rTrigB.Q THEN
            uInfoOne := 16#0003_03F2;                 // 信息级：双请求同拍 A 优先 / Info: simultaneous requests, A first
        END_IF
        IF bEn AND (bReqA OR bReqB) AND (rTrigA.Q OR rTrigB.Q) THEN
            eStep := eMoveAIn;                        // 任一请求沿启动，A 先动 / Any request edge starts, A first
        END_IF
    eMoveAIn:
        IF NOT bEn THEN
            eStep := eIdle;                           // 撤使能回待机 / Disable returns to idle
        ELSIF tonStep.Q THEN
            eStep := eFault;                          // 步超时锁故障 / Step timeout latches fault
            uCodeLatch := 16#0003_03F3;               // 码位：步超时 / Code: step timeout
        ELSIF bPosA AND (NOT bGripA) THEN
            eStep := eFault;                          // 就位未持片反馈矛盾 / In-position without wafer, contradiction
            uCodeLatch := 16#0003_03F5;               // 码位：反馈矛盾 / Code: feedback contradiction
        ELSIF bPosA AND bGripA THEN
            eStep := eMoveBIn;                        // A 就位且持片转 B 进场 / A placed with wafer, B enters
        END_IF
    eMoveBIn:
        IF NOT bEn THEN
            eStep := eIdle;                           // 撤使能回待机 / Disable returns to idle
        ELSIF tonStep.Q THEN
            eStep := eFault;                          // 步超时锁故障 / Step timeout latches fault
            uCodeLatch := 16#0003_03F3;               // 码位：步超时 / Code: step timeout
        ELSIF (NOT bPosA) OR (NOT bGripA) THEN
            eStep := eFault;                          // A 就位窗口非预期丢失 / Unexpected loss of A window
            uCodeLatch := 16#0003_03F5;               // 码位：反馈矛盾 / Code: feedback contradiction
        ELSIF bPosB THEN
            eStep := eARelease;                       // B 就位转 A 释放 / B placed, A releases
        END_IF
    eARelease:
        IF NOT bEn THEN
            eStep := eIdle;                           // 撤使能回待机 / Disable returns to idle
        ELSIF tonStep.Q THEN
            eStep := eFault;                          // 步超时锁故障 / Step timeout latches fault
            uCodeLatch := 16#0003_03F3;               // 码位：步超时 / Code: step timeout
        ELSIF (NOT bPosA) THEN
            eStep := eFault;                          // A 就位窗口非预期丢失 / Unexpected loss of A window
            uCodeLatch := 16#0003_03F5;               // 码位：反馈矛盾 / Code: feedback contradiction
        ELSIF NOT bGripA THEN
            eStep := eWaitGripB;                      // A 释放完成转 B 吸持确认 / A released, wait grip-B
        END_IF
    eWaitGripB:
        IF NOT bEn THEN
            eStep := eIdle;                           // 撤使能回待机 / Disable returns to idle
        ELSIF tonStep.Q THEN
            eStep := eFault;                          // 步超时锁故障 / Step timeout latches fault
            uCodeLatch := 16#0003_03F3;               // 码位：步超时 / Code: step timeout
        ELSIF (NOT bPosA) OR (NOT bPosB) THEN
            eStep := eFault;                          // 就位窗口非预期跳变 / Unexpected position jump
            uCodeLatch := 16#0003_03F5;               // 码位：反馈矛盾 / Code: feedback contradiction
        ELSIF bGripB AND (NOT bGripA) THEN
            eStep := eAExit;                          // B 吸持确认且 A 已释放 / B gripping and A released
        END_IF
    eAExit:
        IF NOT bEn THEN
            eStep := eIdle;                           // 撤使能回待机 / Disable returns to idle
        ELSIF tonStep.Q THEN
            eStep := eFault;                          // 步超时锁故障 / Step timeout latches fault
            uCodeLatch := 16#0003_03F3;               // 码位：步超时 / Code: step timeout
        ELSIF NOT bGripB THEN
            eStep := eFault;                          // B 持片窗口非预期丢失 / Unexpected loss of B wafer
            uCodeLatch := 16#0003_03F5;               // 码位：反馈矛盾 / Code: feedback contradiction
        ELSIF NOT bPosA THEN
            eStep := eBExit;                          // A 撤离完成转 B 撤离 / A exited, B exits
        END_IF
    eBExit:
        IF NOT bEn THEN
            eStep := eIdle;                           // 撤使能回待机 / Disable returns to idle
        ELSIF tonStep.Q THEN
            eStep := eFault;                          // 步超时锁故障 / Step timeout latches fault
            uCodeLatch := 16#0003_03F3;               // 码位：步超时 / Code: step timeout
        ELSIF bPosA THEN
            eStep := eFault;                          // A 非预期重返交接区 / A unexpectedly re-enters zone
            uCodeLatch := 16#0003_03F5;               // 码位：反馈矛盾 / Code: feedback contradiction
        ELSIF NOT bPosB THEN
            eStep := eDone;                           // B 撤离完成转完成态 / B exited, to done
        END_IF
    eDone:
        bDone := TRUE;                                // 完成单拍脉冲 / One-scan done pulse
        eStep := eIdle;                               // 下拍回待机 / Back to idle next scan
    eFault:
        bMoveA := FALSE;                              // 故障态撤 A 放行 / Fault revokes A permit
        bMoveB := FALSE;                              // 故障态撤 B 放行 / Fault revokes B permit
        bDone  := FALSE;                              // 故障态清完成脉冲 / Fault clears done pulse
        IF NOT bEn THEN
            eStep := eIdle;                           // 可达解除路径：撤使能复位 / Reachable release: disable
            uCodeLatch := DL_WHS_ZERO;                // 清锁存码 / Clear latched code
        END_IF
    ELSE
        eStep := eFault;                              // 非法状态兜底 / Illegal state fallback
        uCodeLatch := 16#0003_03F6;                   // 码位：状态非法 / Code: illegal state
END_CASE

// ---- 段 5｜防御断言：双放行同拍为互锁违例（构造上不可达，留档兜底）--------------
IF bMoveA AND bMoveB THEN
    bMoveA := FALSE;                                  // 安全侧撤 A 放行 / Safe side revokes A permit
    bMoveB := FALSE;                                  // 安全侧撤 B 放行 / Safe side revokes B permit
    eStep := eFault;                                  // 互锁违例锁故障 / Interlock violation latches fault
    uCodeLatch := 16#0003_03F4;                       // 码位：互锁违例 / Code: interlock violation
END_IF

// ---- 段 6｜错误码装配：故障锁存回放优先，信息级单拍居次 --------------------------
IF eStep = eFault THEN
    bError   := TRUE;                                 // 故障标志配对（R45）/ Fault flag paired
    uErrorId := uCodeLatch;                           // 故障码锁存回放 / Latched fault code replayed
ELSIF uInfoOne <> DL_WHS_ZERO THEN
    bError   := FALSE;                                // 信息级不置故障 / Info never sets fault
    uErrorId := uInfoOne;                             // 信息级单拍输出 / One-scan info output
    uInfoOne := DL_WHS_ZERO;                          // 发完即清 / Clear after emit
ELSE
    bError   := FALSE;                                // 无错清标志 / Clear fault flag
    uErrorId := DL_WHS_ZERO;                          // 无码 / No code
END_IF
END_FUNCTION_BLOCK

(* ---- FB_DL_WaferMapping.st ---- *)
//==============================================================================
// 功能块：FB_DL_WaferMapping ｜ 中文名称：晶圆花篮（FOUP）Mapping 传感器序列解析
// 所属子库：DL_Device ｜ 版本：v1.0.0 ｜ 兼容：CODESYS V3.5+ / TwinCAT 3 / 汇川 InoProShop
// 功能描述：25 槽在位传感器序列解析 → 逐槽片位图 + 空位/单片/斜插（eCross，
//           相邻槽同时置位）识别 + 在片数统计。序列经 tScanTimeout 稳
//           定判定后才置映射有效（稳定期内任何跳变即重新计时，防抖）。
//           全槽为 0 = 合法空盒，不判故障。只解析与判定，不做机械手
//           动作（取放由上位调度，本件零执行输出）。规格引脚表未提供
//           厚度量测输入，eDouble（双片）判据在本版不可达：枚举保留
//           语义槽，fDoubleThickPct 仅作组态域校验（小于 1.0 判组态非
//           法），待厚度型传感器引脚增补后启用双片判据（主动偏离披露，
//           见修订历史）。
// 开源溯源 (Origin)：道莅原创实现（参考 公开工程惯例 分类与参数域）
// 单位表：槽数[槽] / 槽索引[—] / 厚度倍率[倍] / 扫描稳定超时[ms] / 计数[片]
// 错误码表：16#0003_0196 信息级（存在斜插异常槽但映射整体可判，不置
//           bError）/ 16#0003_0197 信息级（序列含噪跳变提示：同槽连续
//           两拍翻转，不置 bError）/ 16#0003_0372 故障级（在用槽数非
//           法、厚度倍率组态非法或非有限，或全通道同拍跳变（传感器串
//           扰/接线故障），置 bError）/ 16#0003_0373 故障级（片位索引
//           越界：内部访问越界防御槽，正常流程不可达，置 bError）/
//           16#0003_0374 故障级兜底（状态机落 ELSE 或非法状态，置
//           bError 并撤映射）
// 状态机：E_DL_WaferMapState（eIdle=0 / eSampling=10 / eMapped=20 /
//           eFault=99），CASE 含 ELSE 兜底，ELSE 置 0374 并撤映射
//           bMapValid（安全侧：无效映射不得被上位取用）
// 边界行为：① nSlotCount 域 1~25，越界 → 故障 0372；数组访问统一
//           IF nIdx >= 0 AND nIdx < nSlotCount 界检，邻位索引另加
//           nIdx < 25 物理界检（防御槽 0373：正常流程不可达，命中即
//           内部越界防御）；② 全槽 0 = 合法空盒，正常出图，不判故障
//           （空 FOUP 正常工况）；③ 斜插判据：本槽置位且相邻槽（i−1/
//           i+1，双侧边界防护）也置位 → 两槽均判 eCross；④ 全通道同
//           拍跳变（上一拍全 0 本拍全 1 或反之）→ 故障 0372（传感器
//           串扰/接线故障），映射撤，故障锁存待 bReset 或失能恢复；
//           ⑤ 异常但可判（有斜插槽）→ 信息 0196；同槽连续两拍翻转 →
//           信息 0197（含噪跳变提示，优先级低于 0196 不覆盖）；⑥ 厚
//           度倍率组态非法（小于 1.0）或非有限 → 故障 0372（数据不可
//           信同语义，复用组态槽不新占码位）；⑦ 失能 → 撤映射、计数
//           清零；⑧ 序列稳定（tScanTimeout 内无跳变）才置 bMapValid，
//           稳定定时器经跳变「断输入一拍」重启（R40 家族）；⑨ 上电
//           首拍 bMapValid := FALSE。
// 修订历史：v1.0.0 2026-11-17 首版（R25 派单 · §4.7）
//==============================================================================
(*------------------------------------------------------------------------------
 * 枚举: E_DL_SlotKind / E_DL_WaferMapState（归属 DL_Device，与 FB_DL_WaferMapping 同文件）
 *----------------------------------------------------------------------------*)
TYPE E_DL_SlotKind :
(
    eEmpty   := 0,   // 空位：传感器未置位 / Empty: sensor off
    eSingle  := 1,   // 单片：本槽置位且相邻无片 / Single: occupied with no occupied neighbor
    eDouble  := 2,   // 双片（斜插厚度型）：本版不可达，语义保留槽 / Double wafer: unreachable this version, semantic slot reserved
    eCross   := 3,   // 斜插：本槽与相邻槽同时置位 / Crossed wafer: occupied with an occupied neighbor
    eUnknown := 4    // 未知：本版 BOOL 序列不可达，语义保留槽 / Unknown: unreachable with BOOL sequence this version
);
END_TYPE
TYPE E_DL_WaferMapState :
(
    eIdle     := 0,   // 失能/待机：映射撤、计数清零 / Idle: mapping withdrawn, counts zeroed
    eSampling := 10,  // 采样中：序列未稳定，映射暂不可取用 / Sampling: sequence not stable, mapping not usable yet
    eMapped   := 20,  // 映射有效：序列稳定期满，结果可取用 / Mapped: stable period elapsed, results usable
    eFault    := 99   // 故障兜底态：组态非法/串扰/非法状态，映射撤 / Fault fallback, mapping withdrawn
);
END_TYPE
FUNCTION_BLOCK FB_DL_WaferMapping
VAR_INPUT
    abSlotSensor  : ARRAY[0..24] OF BOOL;      // 逐槽在位信号，长度固定 25 [—] / Per-slot wafer-present signals, fixed length 25
    nSlotCount    : INT := 25;                 // 在用槽数 [槽]，1~25 / Slots in use, 1~25
    fDoubleThickPct : LREAL := 1.5;            // 厚度倍率判双片 [倍]，本版仅做组态域校验 / Thickness ratio for double detection, config-validated only this version
    tScanTimeout  : TIME := T#10S;             // 扫描稳定超时 [ms]，稳定期满映射生效 / Scan stability timeout [ms]
    bEnable       : BOOL;                      // 总使能 / Master enable
    bReset        : BOOL;                      // 复位，上升沿清状态与计数 / Reset, rising edge clears state and counters
END_VAR
VAR_OUTPUT
    abSlotOccupied : ARRAY[0..24] OF BOOL;     // 逐槽在位映射（稳定期内可取用）/ Per-slot occupancy map, usable while stable
    aeSlotKind    : ARRAY[0..24] OF E_DL_SlotKind;  // 逐槽片型判定 / Per-slot wafer kind verdict
    nOccupiedCount : INT;                      // 在片数 [片] / Occupied slot count
    bMapValid     : BOOL;                      // 映射有效标志：序列稳定期满且无故障 / Mapping valid: stable period elapsed and no fault
    bAnyAnomaly   : BOOL;                      // 存在异常槽（斜插等）但映射整体可判 / Any anomalous slot while map still judgeable
    nAnomalyCount : INT;                       // 异常槽数 [槽] / Anomalous slot count
    eErr          : UDINT;                     // 错误码，0 = 无错，码位 16#0003_0196 起信息级、16#0003_0372 起故障级（分带见错误码表） / Error code, 0 = no error, band info/fault per the code table
    bError        : BOOL;                      // 故障级标志，仅故障级错误置位 / Fault-class flag, set only on fault-level codes
    bValid        : BOOL;                      // 判定数据可用标志，失能/故障闸显式 FALSE / Verdict usable flag, explicit FALSE on disable/fault gates
    eState        : E_DL_WaferMapState;        // 主状态机当前状态 / Current state of the main state machine
END_VAR
VAR
    fbReset       : R_TRIG;                    // 复位上升沿检测实例 / Reset rising edge detector
    fbStableT     : TON;                       // 序列稳定定时器（跳变断输入一拍重启）/ Sequence stability timer, kicked on change
    bStableKick   : BOOL;                      // 稳定定时器断输入一拍标志（R40 家族）/ Stability timer one-scan kick flag
    abPrev        : ARRAY[0..24] OF BOOL;      // 上一拍逐槽快照（跳变检测）/ Previous-scan per-slot snapshot for change detection
    abChg         : ARRAY[0..24] OF BOOL;      // 本拍逐槽跳变标志 / Per-slot change flag this scan
    abChgPrev     : ARRAY[0..24] OF BOOL;      // 上一拍逐槽跳变标志（含噪翻转检测）/ Previous-scan change flags for flap detection
    nChgCount     : INT;                       // 本拍跳变槽总数 [槽] / Total changed slots this scan
    bAllSameNow   : BOOL;                      // 本拍全槽同值判据 / All slots equal this scan
    bAllValNow    : BOOL;                      // 本拍全槽同值时的值 / The common value when all equal this scan
    bAllSamePrev  : BOOL;                      // 上一拍全槽同值判据 / All slots equal previous scan
    bAllValPrev   : BOOL;                      // 上一拍全槽同值时的值 / The common value when all equal previous scan
    bCrossJump    : BOOL;                      // 全通道同拍跳变（串扰判据）/ Whole-array same-scan jump (crosstalk criterion)
    bNoiseFlap    : BOOL;                      // 含噪跳变：同槽连续两拍翻转 / Noisy flap: same slot toggling two scans in a row
    uIdx          : INT;                       // 槽循环索引 [—] / Slot loop index
    nNb           : INT;                       // 邻位槽索引 [—] / Neighbor slot index
    bNbOccupied   : BOOL;                      // 邻位在位判据（双侧边界防护）/ Neighbor occupied predicate, double-side bounded
    nOccCount     : INT;                       // 在片数暂存 [片] / Occupied count staging
    nAnomCount    : INT;                       // 异常槽数暂存 [槽] / Anomaly count staging
    bPrevValid    : BOOL;                      // 上一拍快照有效标志（首拍跳变检测屏蔽）/ Previous snapshot valid, first-scan jump masked
END_VAR
VAR CONSTANT
    DL_WMAP_CODE_INFO_1 : UDINT := 16#0003_0196;  // 信息级槽 1（异常但映射可判） / info slot 1
    DL_WMAP_CODE_INFO_2 : UDINT := 16#0003_0197;  // 信息级槽 2（序列含噪跳变提示） / info slot 2
    DL_WMAP_CODE_FLT_1  : UDINT := 16#0003_0372;  // 故障级槽 1（槽数非法或串扰跳变） / fault slot 1
    DL_WMAP_CODE_FLT_2  : UDINT := 16#0003_0373;  // 故障级槽 2（片位索引越界防御） / fault slot 2
    DL_WMAP_CODE_FLT_3  : UDINT := 16#0003_0374;  // 故障级槽 3（非法状态兜底） / fault slot 3, illegal-state fallback
    DL_WM_SLOT_MAX : INT := 25;                // 槽数硬上限 [槽]，数组物理长度 / Slot hard ceiling, array physical length
    DL_WM_ZERO     : INT := 0;                 // 零值常量，避免裸字面量 [—] / Zero constant, avoids a bare literal
    DL_WM_ONE      : INT := 1;                 // 一值常量，避免裸字面量 [—] / One constant, avoids a bare literal
    DL_WM_RATIO_MIN : LREAL := 1.0;            // 厚度倍率组态下限 [倍] / Thickness ratio config floor
    DL_WM_INF      : LREAL := 1.7976931348623157E308;  // LREAL 幅值上限，Inf 判据 / LREAL magnitude ceiling, Inf criterion
END_VAR

(*------------------------------------------------------------------------------
 * 段 1｜无条件刷新区（红线 5）：复位沿与稳定定时器在任何分支之外周期调用
 *----------------------------------------------------------------------------*)
fbReset(CLK := bReset);                        // 复位沿检测无条件刷新 / reset edge refreshed unconditionally
fbStableT(IN := bEnable AND (NOT bStableKick),  // 稳定计时：使能且本拍无跳变断输入（R40 家族）/ stability timing, kicked on any change
          PT := tScanTimeout);                 // 稳定期门槛 / stability threshold
bStableKick := FALSE;                          // kick 标志单拍自清（跳变时由采样段重置位）/ kick self-clears, re-set on change

(*------------------------------------------------------------------------------
 * 段 2｜复位沿处理（改写置于沿后，防吞沿 R39）
 *----------------------------------------------------------------------------*)
IF fbReset.Q THEN
    eState     := E_DL_WaferMapState.eIdle;
    eErr       := 16#0000_0000;                // 复位清码 / reset clears code
    bError     := FALSE;                       // 复位清故障 / reset clears fault
    bMapValid  := FALSE;                       // 映射撤 / mapping withdrawn
    bAnyAnomaly := FALSE;                      // 异常标志清 / anomaly flag cleared
    nAnomalyCount := DL_WM_ZERO;               // 异常计数清零 / anomaly count zeroed
    nOccupiedCount := DL_WM_ZERO;              // 在片数清零 / occupied count zeroed
    bPrevValid := FALSE;                       // 首拍跳变检测重新屏蔽 / first-scan jump masked again
    FOR uIdx := 0 TO 24 DO
        abPrev[uIdx] := FALSE;                 // 上一拍快照清零 / previous snapshot zeroed
        abChg[uIdx] := FALSE;                  // 跳变标志清零 / change flags zeroed
        abChgPrev[uIdx] := FALSE;              // 上一拍跳变标志清零 / previous change flags zeroed
        abSlotOccupied[uIdx] := FALSE;         // 映射输出清零 / occupancy outputs zeroed
        aeSlotKind[uIdx] := E_DL_SlotKind.eEmpty;  // 片型输出清空位 / kind outputs to empty
    END_FOR
END_IF

(*------------------------------------------------------------------------------
 * 段 3｜组态与非有限闸（槽数域 / 厚度倍率域，非有限复用 0372 不新占码位）
 *----------------------------------------------------------------------------*)
IF (nSlotCount < DL_WM_ONE) OR (nSlotCount > DL_WM_SLOT_MAX)
   OR (fDoubleThickPct <> fDoubleThickPct) OR (ABS(fDoubleThickPct) >= DL_WM_INF)
   OR (fDoubleThickPct < DL_WM_RATIO_MIN) THEN
    eState    := E_DL_WaferMapState.eFault;
    eErr      := DL_WMAP_CODE_FLT_1;               // 故障级：槽数非法或厚度倍率组态非法/非有限 / fault: slot count or ratio config invalid
    bError    := TRUE;                         // 故障级必置 bError（R45 配对）/ fault-class pairs with bError
    bValid    := FALSE;                        // 输出不可用 / outputs unusable
    bMapValid := FALSE;                        // 映射撤（安全侧）/ mapping withdrawn, safe side
    bAnyAnomaly := FALSE;                      // 故障态不判异常 / anomaly not judged in fault
    nAnomalyCount := DL_WM_ZERO;               // 异常计数清零 / anomaly count zeroed
    nOccupiedCount := DL_WM_ZERO;              // 在片数清零 / occupied count zeroed
    fbStableT(IN := FALSE, PT := tScanTimeout);  // 稳定定时器断输入（无条件调用保持）/ stability timer input broken, still called
    RETURN;
END_IF

(*------------------------------------------------------------------------------
 * 段 4｜逐槽界检快照对比：跳变标志、全同判据、串扰判据（防御槽 0373）
 *----------------------------------------------------------------------------*)
nChgCount := DL_WM_ZERO;                       // 跳变计数清零 / change count zeroed
bAllSameNow := TRUE;                           // 全同判据种子 / all-equal predicate seed
bAllValNow := abSlotSensor[0];                 // 全同参考值种子 / all-equal reference seed
FOR uIdx := 0 TO 24 DO
    IF (uIdx < DL_WM_ZERO) OR (uIdx >= DL_WM_SLOT_MAX) THEN
        eState := E_DL_WaferMapState.eFault;   // 片位索引越界（内部防御，正常不可达）/ slot index out of bounds, defensive
        eErr := DL_WMAP_CODE_FLT_2;                // 故障级：片位索引越界 / fault: slot index out of bounds
        bError := TRUE;                        // 故障级必置 bError / fault-class pairs with bError
        bValid := FALSE;                       // 输出不可用 / outputs unusable
        bMapValid := FALSE;                    // 映射撤（安全侧）/ mapping withdrawn, safe side
        fbStableT(IN := FALSE, PT := tScanTimeout);  // 稳定定时器断输入（无条件调用保持）/ stability timer input broken
        RETURN;
    END_IF
    IF abSlotSensor[uIdx] <> bAllValNow THEN
        bAllSameNow := FALSE;                  // 有异值即非全同 / any differing value breaks all-equal
    END_IF
    abChg[uIdx] := bPrevValid AND (abSlotSensor[uIdx] <> abPrev[uIdx]);  // 逐槽跳变标志（首拍屏蔽）/ per-slot change flag, masked on first scan
    IF abChg[uIdx] THEN
        nChgCount := nChgCount + DL_WM_ONE;    // 跳变槽计数 / count changed slot
        bStableKick := TRUE;                   // 任一跳变：稳定定时器断输入一拍重启 / any change kicks the stability timer
    END_IF
END_FOR
bCrossJump := bPrevValid AND bAllSameNow AND bAllSamePrev AND (bAllValNow <> bAllValPrev);  // 全通道同拍跳变判据 / whole-array jump predicate
bNoiseFlap := FALSE;                           // 含噪判据复位 / noise criterion reset
FOR uIdx := 0 TO 24 DO
    IF abChg[uIdx] AND abChgPrev[uIdx] THEN
        bNoiseFlap := TRUE;                    // 同槽连续两拍翻转 → 信息 0197 / same slot toggling two scans in a row
    END_IF
END_FOR

(*------------------------------------------------------------------------------
 * 段 5｜分类与计数：逐槽界检 + 邻位双侧边界防护，斜插两槽均判 eCross
 *----------------------------------------------------------------------------*)
nOccCount := DL_WM_ZERO;                       // 在片数清零 / occupied count zeroed
nAnomCount := DL_WM_ZERO;                      // 异常数清零 / anomaly count zeroed
FOR uIdx := 0 TO 24 DO
    IF uIdx < nSlotCount THEN
        abSlotOccupied[uIdx] := abSlotSensor[uIdx];  // 在用槽：照抄传感器 / in-use slot: copy sensor
        IF abSlotSensor[uIdx] THEN
            bNbOccupied := FALSE;              // 邻位在位判据复位 / neighbor predicate reset
            nNb := uIdx - DL_WM_ONE;           // 左邻索引 / left neighbor index
            IF (nNb >= DL_WM_ZERO) AND (nNb < nSlotCount) AND (nNb < DL_WM_SLOT_MAX) THEN
                IF abSlotSensor[nNb] THEN
                    bNbOccupied := TRUE;       // 左邻在位 / left neighbor occupied
                END_IF
            END_IF
            nNb := uIdx + DL_WM_ONE;           // 右邻索引 / right neighbor index
            IF (nNb >= DL_WM_ZERO) AND (nNb < nSlotCount) AND (nNb < DL_WM_SLOT_MAX) THEN
                IF abSlotSensor[nNb] THEN
                    bNbOccupied := TRUE;       // 右邻在位 / right neighbor occupied
                END_IF
            END_IF
            IF bNbOccupied THEN
                aeSlotKind[uIdx] := E_DL_SlotKind.eCross;  // 斜插：相邻同时置位 / crossed: adjacent occupied
                nAnomCount := nAnomCount + DL_WM_ONE;      // 异常槽计数 / count anomalous slot
            ELSE
                aeSlotKind[uIdx] := E_DL_SlotKind.eSingle; // 单片：邻位无片 / single: no occupied neighbor
            END_IF
            nOccCount := nOccCount + DL_WM_ONE;        // 在片计数 / count occupied slot
        ELSE
            aeSlotKind[uIdx] := E_DL_SlotKind.eEmpty;  // 空位 / empty
        END_IF
    ELSE
        abSlotOccupied[uIdx] := FALSE;         // 超出在用槽数：按空位出图 / beyond in-use count: mapped empty
        aeSlotKind[uIdx] := E_DL_SlotKind.eEmpty;  // 片型空位 / kind empty
    END_IF
END_FOR
nOccupiedCount := nOccCount;                   // 在片数出口 / occupied count output
nAnomalyCount := nAnomCount;                   // 异常数出口 / anomaly count output
bAnyAnomaly := nAnomCount > DL_WM_ZERO;        // 异常标志 / anomaly flag

(*------------------------------------------------------------------------------
 * 段 6｜历史快照滚动：本拍值与跳变标志存为上一拍（供下拍对比）
 *----------------------------------------------------------------------------*)
FOR uIdx := 0 TO 24 DO
    abPrev[uIdx] := abSlotSensor[uIdx];        // 滚动值快照 / roll value snapshot
    abChgPrev[uIdx] := abChg[uIdx];            // 滚动跳变快照 / roll change snapshot
END_FOR
bPrevValid := TRUE;                            // 快照有效 / snapshot valid
bAllSamePrev := bAllSameNow;                   // 滚动全同判据 / roll all-equal predicate
bAllValPrev := bAllValNow;                     // 滚动全同参考值 / roll all-equal reference

(*------------------------------------------------------------------------------
 * 段 7｜状态机：CASE 含 ELSE 兜底（非法状态 → 0374 + 撤映射，安全侧）
 *----------------------------------------------------------------------------*)
CASE eState OF

    E_DL_WaferMapState.eIdle:
        bValid := FALSE;                       // 失能闸显式不可用（R72）/ explicit FALSE on disable gate
        bMapValid := FALSE;                    // 映射撤 / mapping withdrawn
        eErr := 16#0000_0000;                  // 待机无错 / no error in idle
        bError := FALSE;                       // 待机无故障 / no fault in idle
        IF bEnable THEN
            eState := E_DL_WaferMapState.eSampling;    // 使能进采样 / enable enters sampling
            bPrevValid := FALSE;               // 重新首拍屏蔽跳变检测 / mask jump detection on fresh start
            bStableKick := TRUE;               // 稳定定时器重启 / stability timer restarted
        END_IF

    E_DL_WaferMapState.eSampling:
        bValid := TRUE;                        // 采样态判定数据可用（bMapValid 仍假）/ verdict usable in sampling, map still not valid
        bMapValid := FALSE;                    // 序列未稳定，映射暂不可取用 / sequence not stable, mapping not usable
        IF NOT bEnable THEN
            eState := E_DL_WaferMapState.eIdle;        // 失能回待机 / disable returns to idle
            bValid := FALSE;                   // 失能闸显式不可用 / explicit FALSE on disable gate
        ELSIF bCrossJump THEN
            eState := E_DL_WaferMapState.eFault;       // 全通道同拍跳变进故障（锁存待复位）/ whole-array jump enters fault, latched
            eErr := DL_WMAP_CODE_FLT_1;            // 故障级：传感器串扰/接线故障 / fault: crosstalk or wiring
            bError := TRUE;                    // 故障级必置 bError / fault-class pairs with bError
            bMapValid := FALSE;                // 映射撤（安全侧）/ mapping withdrawn, safe side
        ELSIF fbStableT.Q THEN
            eState := E_DL_WaferMapState.eMapped;      // 稳定期满映射生效 / stability elapsed, mapping valid
        END_IF

    E_DL_WaferMapState.eMapped:
        bValid := TRUE;                        // 映射态判定数据可用 / verdict usable in mapped
        bMapValid := TRUE;                     // 映射有效 / mapping valid
        IF NOT bEnable THEN
            eState := E_DL_WaferMapState.eIdle;
            bValid := FALSE;                   // 失能闸显式不可用 / explicit FALSE on disable gate
            bMapValid := FALSE;                // 映射撤 / mapping withdrawn
        ELSIF bCrossJump THEN
            eState := E_DL_WaferMapState.eFault;       // 全通道同拍跳变进故障（锁存待复位）/ whole-array jump enters fault, latched
            eErr := DL_WMAP_CODE_FLT_1;
            bError := TRUE;
            bMapValid := FALSE;                // 映射撤（安全侧）/ mapping withdrawn, safe side
        ELSIF nChgCount > DL_WM_ZERO THEN
            eState := E_DL_WaferMapState.eSampling;    // 稳定期内出现跳变回采样 / change during stable period returns to sampling
            bMapValid := FALSE;                // 映射暂撤 / mapping withdrawn temporarily
        END_IF

    E_DL_WaferMapState.eFault:
        bValid := FALSE;                       // 故障闸显式不可用 / explicit FALSE on fault gate
        bMapValid := FALSE;                    // 映射撤（安全侧）/ mapping withdrawn, safe side
        eErr := DL_WMAP_CODE_FLT_1;                // 故障级保持（串扰或组态，见进入路径）/ fault held
        bError := TRUE;                        // 故障级必置 bError / fault-class pairs with bError
        IF NOT bEnable THEN
            eState := E_DL_WaferMapState.eIdle;        // 仅失能解锁（串扰故障锁存，见边界行为④；bReset 走段 2 路径）/ only disable unlocks, crosstalk latched, reset via section 2
        END_IF

    ELSE
        eState := E_DL_WaferMapState.eFault;   // 非法状态兜底 / illegal-state fallback
        eErr := DL_WMAP_CODE_FLT_3;                // 故障级兜底：非法状态 / fault fallback: illegal state
        bError := TRUE;                        // 故障级必置 bError / fault-class pairs with bError
        bValid := FALSE;                       // 输出不可用 / outputs unusable
        bMapValid := FALSE;                    // 映射撤（安全侧，无效映射不得被取用）/ mapping withdrawn, safe side
END_CASE

(*------------------------------------------------------------------------------
 * 段 8｜信息级收口：0196 异常可判 与 0197 含噪提示（均不置 bError）
 *----------------------------------------------------------------------------*)
IF bAnyAnomaly AND (eState = E_DL_WaferMapState.eMapped) THEN
    eErr := DL_WMAP_CODE_INFO_1;               // 信息级：存在斜插异常但映射整体可判 / info: anomaly present, map judgeable
    bError := FALSE;                           // 信息级不置 bError / info never raises bError
END_IF
IF bNoiseFlap AND (eState = E_DL_WaferMapState.eSampling OR eState = E_DL_WaferMapState.eMapped) THEN
    eErr := DL_WMAP_CODE_INFO_2;               // 信息级：同槽连续两拍翻转含噪提示 / info: noisy same-slot flap
    bError := FALSE;                           // 信息级不置 bError / info never raises bError
END_IF
END_FUNCTION_BLOCK
